(* IEC 61131-3 sources: RootPLC/conformance/cases/statements, 14 files *)

(* ---- err_duplicate_argument.st ---- *)
(* spec: [statements.call]
   expect: error RP0302 *)
FUNCTION_BLOCK FB_Lamp
VAR_INPUT
    lit : BOOL;
END_VAR
END_FUNCTION_BLOCK

PROGRAM P
VAR
    lamp : FB_Lamp;
END_VAR
lamp(lit := TRUE, LIT := FALSE);
END_PROGRAM

(* ---- ok_case_timer_reset.st ---- *)
(* spec: [statements.case.timer]
   expect: ok *)
(* Three ways to time a step without RP0304. *)
FUNCTION_BLOCK FB_Steps
VAR_INPUT go : BOOL; done : BOOL; END_VAR
VAR
    a : INT;
    b : INT;
    c : INT;
    tA : TON;
    tB : TON;
    tC : TON;
END_VAR
(* every path that leaves the step stops the timer first *)
CASE a OF
    0:
        IF go THEN a := 1; END_IF;
    1:
        tA(IN := TRUE, PT := T#5s);
        IF done OR tA.Q THEN
            tA(IN := FALSE);
            a := 0;
        END_IF;
END_CASE;
(* reset in the step before: cleared before re-entry *)
CASE b OF
    0:
        tB(IN := FALSE);
        IF go THEN b := 1; END_IF;
    1:
        tB(IN := TRUE, PT := T#5s);
        IF tB.Q THEN b := 0; END_IF;
END_CASE;
(* called every cycle outside the CASE with the step condition *)
tC(IN := c = 1, PT := T#5s);
CASE c OF
    0:
        IF go THEN c := 1; END_IF;
    1:
        IF tC.Q THEN c := 0; END_IF;
END_CASE;
END_FUNCTION_BLOCK

(* ---- warn_call_empty_input.st ---- *)
(* spec: [statements.call] [scope.vendor-forms]
   expect: warning RP0118 RP0134
   run: PRG_Main cycles=1
   assert: k = 4
   assert: n = 4 *)
FUNCTION_BLOCK FB_Store
VAR_INPUT
    v : INT;
    flag : BOOL := TRUE;
END_VAR
VAR_OUTPUT
    k : INT;
END_VAR
k := v;
END_FUNCTION_BLOCK

FUNCTION F_Len : INT
VAR_INPUT
    s : REFERENCE TO STRING;
END_VAR
F_Len := LEN(s);
END_FUNCTION

PROGRAM PRG_Main
VAR
    f : FB_Store;
    k, n : INT;
    txt : STRING := 'abcd';
END_VAR
f(v := 4, flag :=, );
k := f.k;
n := F_Len(txt);
END_PROGRAM

(* ---- warn_call_empty_output.st ---- *)
(* spec: [statements.call] [scope.vendor-forms]
   expect: warning RP0134
   run: PRG_Main cycles=1
   assert: n = 4 *)
FUNCTION_BLOCK FB_Count
VAR_INPUT
    k : INT;
END_VAR
VAR_OUTPUT
    Done : BOOL;
    Count : INT;
END_VAR
Done := TRUE;
Count := k;
END_FUNCTION_BLOCK

PROGRAM PRG_Main
VAR
    f : FB_Count;
    n : INT;
END_VAR
f(k := 4, Done =>, Count => n);
END_PROGRAM

(* ---- warn_case_timer_left_running.st ---- *)
(* spec: [statements.case.timer]
   expect: warning RP0304 *)
(* The timeout path leaves step 1 while tTimeout still has IN = TRUE: after
   Reset, the next homing faults on its first call (found in real code). *)
FUNCTION_BLOCK FB_Home
VAR_INPUT start : BOOL; atHome : BOOL; reset : BOOL; END_VAR
VAR_OUTPUT move : BOOL; fault : BOOL; END_VAR
VAR nStep : INT; tTimeout : TON; END_VAR
CASE nStep OF
    0:
        IF start THEN
            nStep := 1;
        END_IF;
    1:
        tTimeout(IN := TRUE, PT := T#10s);
        IF atHome THEN
            tTimeout(IN := FALSE);
            nStep := 2;
        ELSIF tTimeout.Q THEN
            nStep := 99;
        END_IF;
    2:
        IF reset THEN
            nStep := 0;
        END_IF;
    99:
        IF reset THEN
            nStep := 0;
        END_IF;
END_CASE;
move := nStep = 1;
fault := nStep = 99;
END_FUNCTION_BLOCK

(* ---- err_missing_semicolon.st ---- *)
(* spec: [statements.terminator]
   expect: error RP0301 *)
PROGRAM PRG_Main
VAR
    x : INT;
END_VAR
x := 1
END_PROGRAM

(* ---- ok_case.st ---- *)
(* spec: [statements.case]
   expect: ok
   run: PRG_Main cycles=1
   assert: r = 2 *)
PROGRAM PRG_Main
VAR
    n : INT := 7;
    r : INT;
END_VAR
CASE n OF
    1, 2:
        r := 1;
    3..9:
        r := 2;
ELSE
    r := 0;
END_CASE;
END_PROGRAM

(* ---- ok_if_else.st ---- *)
(* spec: [statements.if]
   expect: ok
   run: PRG_Main cycles=1
   assert: y = 2 *)
PROGRAM PRG_Main
VAR
    x : INT := 5;
    y : INT;
END_VAR
IF x > 3 THEN
    y := 2;
ELSE
    y := 1;
END_IF;
END_PROGRAM

(* ---- ok_loops.st ---- *)
(* spec: [statements.for] [statements.while] [statements.repeat] [statements.control] [scope.iec]
   expect: ok
   run: PRG_Main cycles=1
   assert: s = 31
   assert: w = 3
   assert: k = 6 *)
PROGRAM PRG_Main
VAR
    i, s, w, k : INT;
END_VAR
FOR i := 1 TO 10 BY 1 DO
    IF i = 5 THEN
        CONTINUE;
    END_IF;
    IF i > 8 THEN
        EXIT;
    END_IF;
    s := s + i;
END_FOR;
WHILE w < 3 DO
    w := w + 1;
END_WHILE;
REPEAT
    k := k + 2;
UNTIL k >= 6
END_REPEAT;
RETURN;
END_PROGRAM

(* ---- ok_precedence.st ---- *)
(* spec: [statements.expression.precedence] [statements.expression.access] [syntax.lossless]
   expect: ok
   run: PRG_Main cycles=1
   assert: a = 50
   assert: b = TRUE
   assert: c = TRUE
   assert: d = 4
   assert: arr[1, 1] = 50
   assert: p.x = 5 *)
TYPE Point : STRUCT x : INT; END_STRUCT; END_TYPE

PROGRAM PRG_Main
VAR
    a : INT;
    b, c : BOOL;
    d : INT;
    arr : ARRAY[0..1, 0..1] OF INT;
    p : Point;
    r : REF_TO Point;
END_VAR
a := 2 + 3 * 4 ** 2;      // 50
b := NOT FALSE OR FALSE;  (* TRUE *)
c := 1 + 2 = 3;
d := -2 ** 2;             /* 4 */
arr[1, 1] := a;
r := REF(p);
r^.x := 5;
END_PROGRAM

(* ---- warn_case_enum_dot.st ---- *)
(* spec: [types.derived.enum]
   expect: warning RP0122
   run: PRG_Main cycles=1
   assert: x = 2 *)
TYPE E_Step : (Idle, Moving, Done); END_TYPE

PROGRAM PRG_Main
VAR
    s : E_Step := E_Step#Moving;
    x : INT;
END_VAR
CASE s OF
    E_Step.Idle:
        x := 1;
    E_Step.Moving, E_Step.Done:
        x := 2;
ELSE
    x := 3;
END_CASE;
END_PROGRAM

(* ---- warn_chained_assign.st ---- *)
(* spec: [statements.assignment.chain]
   expect: warning RP0125
   run: PRG_Main cycles=1
   assert: a = 7
   assert: b = 7
   assert: c = 7 *)
PROGRAM PRG_Main
VAR
    a, b, c : INT;
END_VAR
a := b := c := 7;
END_PROGRAM

(* ---- warn_for_element_control.st ---- *)
(* spec: [statements.for] [scope.vendor-forms]
   expect: warning RP0134
   run: PRG_Main cycles=1
   assert: sum = 10 *)
PROGRAM PRG_Main
VAR
    idx : ARRAY[1..2] OF INT;
    sum : INT;
END_VAR
FOR idx[1] := 1 TO 4 DO
    sum := sum + idx[1];
END_FOR;
END_PROGRAM

(* ---- warn_set_reset_assign.st ---- *)
(* spec: [statements.assignment.set-reset]
   expect: warning RP0123
   run: PRG_Main cycles=1
   assert: a = TRUE
   assert: b = FALSE
   assert: c = TRUE *)
PROGRAM PRG_Main
VAR
    a : BOOL;
    b : BOOL := TRUE;
    c : BOOL := TRUE;
    go : BOOL := TRUE;
END_VAR
a S= go;
b R= go;
c R= NOT go;
END_PROGRAM
